Staubli VAL3: initContainer.pgx

public program initContainer(utContainer& x_utContainer[], string x_sPage, string x_sId, bool x_bVisibility)
begin
  x_utContainer.Common.sPage=x_sPage
  x_utContainer.Common.sID=x_sId
  userPageBind(x_utContainer.Common.sPage,x_utContainer.Common.sID,"src",x_utContainer.Common.sSource,1,"r")
  userPageBind(x_utContainer.Common.sPage,x_utContainer.Common.sID,"style.visibility",x_utContainer.Appearance.bVisibility,1,"r")
  //
  x_utContainer.Appearance.bVisibility=x_bVisibility
end
